Fanuc KAREL source: kx00027.compact.KL

PROGRAM KX00027
%STACKSIZE=1000
%PRIORITY=65535
%NOLOCKGROUP
VAR
I : INTEGER
J : INTEGER
B : BOOLEAN
F : FILE
S : STRING[80]
P : XYZWPR
BEGIN
I=1
END KX00027
